(* IEC 61131-3 sources: plc-st-coding-agent/progress/evidence/f14_p1_20261111b/jobs/custom_deepseek-v4pro (part 2) *)

(* ---- self-hard-05.candidate_02.st ---- *)
FUNCTION_BLOCK FB
VAR_INPUT
    runRequest : BOOL;
    flameOK : BOOL;
    o2Valid : BOOL;
    o2PV : REAL;
    baseAir : REAL;
    resetBtn : BOOL;
END_VAR
VAR_OUTPUT
    fuelPermit : BOOL;
    trimEnable : BOOL;
    airTrim : REAL;
    airCommand : REAL;
    tripLatched : BOOL;
    o2Fault : BOOL;
END_VAR
VAR
    tripState : BOOL := FALSE;   (* internal trip memory *)
    prevReset : BOOL := FALSE;   (* previous cycle reset button state *)
    resetRising : BOOL;          (* reset rising edge flag *)
    rawTrim : REAL;              (* unclamped oxygen trim *)
END_VAR
BEGIN
    (* 1. Analyzer fault detection *)
    o2Fault := (NOT o2Valid) OR (o2PV < 0.0) OR (o2PV > 21.0);

    (* 2. Reset button rising edge detection *)
    resetRising := resetBtn AND (NOT prevReset);

    (* 3. Trip state update (immediate set, self-holding with edge-clear) *)
    IF (runRequest AND (NOT flameOK)) THEN
        tripState := TRUE;
    ELSIF (tripState AND resetRising AND (NOT runRequest) AND (NOT flameOK)) THEN
        tripState := FALSE;
    END_IF;

    (* 4. Output latched trip *)
    tripLatched := tripState;

    (* 5. Fuel permit *)
    fuelPermit := runRequest AND flameOK AND (NOT tripLatched);

    (* 6. Oxygen trim enable *)
    trimEnable := fuelPermit AND (NOT o2Fault);

    (* 7. Oxygen trim calculation *)
    IF trimEnable THEN
        rawTrim := 2.0 * (2.0 - o2PV);
        IF rawTrim < -10.0 THEN
            airTrim := -10.0;
        ELSIF rawTrim > 10.0 THEN
            airTrim := 10.0;
        ELSE
            airTrim := rawTrim;
        END_IF;
    ELSE
        airTrim := 0.0;
    END_IF;

    (* 8. Air command calculation *)
    IF fuelPermit THEN
        airCommand := baseAir + airTrim;
        IF airCommand < 0.0 THEN
            airCommand := 0.0;
        ELSIF airCommand > 100.0 THEN
            airCommand := 100.0;
        END_IF;
    ELSE
        airCommand := 0.0;
    END_IF;

    (* 9. Store reset button state for next cycle edge detection *)
    prevReset := resetBtn;
END_FUNCTION_BLOCK

(* ---- self-hard-06.candidate_01.st ---- *)
FUNCTION_BLOCK FB
VAR_INPUT
    runRequest : BOOL;
    pressure : REAL;
    pressureValid : BOOL;
    fuelFlow : REAL;
    steamFlow : REAL;
    outletCmd : INT;
    outletFeedback : INT;
    resetBtn : BOOL;
END_VAR
VAR_OUTPUT
    tripLatched : BOOL;
    fuelPermit : BOOL;
    currentCauseMask : WORD;
    latchedCauseMask : WORD;
    diagnosticActive : BOOL;
END_VAR
VAR
    stallCount : INT := 0;          (* 连续卡滞计数 *)
    prevResetBtn : BOOL := FALSE;   (* 上一周期复位按钮 *)
    risingReset : BOOL;
    condStall : BOOL;
    newTripLatched : BOOL;
END_VAR

(* 复位按钮上升沿检测 *)
risingReset := resetBtn AND NOT prevResetBtn;

(* 计算本拍诊断线索 currentCauseMask *)
currentCauseMask := 0;

IF NOT runRequest THEN
    currentCauseMask := 0;
    stallCount := 0;
ELSIF NOT pressureValid THEN
    currentCauseMask := 1;          (* bit0: 变送器失效 *)
    stallCount := 0;
ELSE
    (* runRequest AND pressureValid *)
    IF pressure < 4500.0 THEN
        currentCauseMask := 0;
        stallCount := 0;
    ELSE
        (* 超压工况: pressure >= 4500.0 *)
        condStall := (outletCmd >= 50) AND (outletFeedback <= 10);
        IF condStall THEN
            stallCount := stallCount + 1;
        ELSE
            stallCount := 0;
        END_IF

        (* bit1: 减温减压阀卡滞，连续3拍 *)
        IF stallCount >= 3 THEN
            currentCauseMask := currentCauseMask OR 16#0002;
        END_IF

        (* bit2: 燃烧过剩 *)
        IF (fuelFlow >= 4.0) AND (steamFlow <= 10.0) THEN
            currentCauseMask := currentCauseMask OR 16#0004;
        END_IF

        (* bit3: 未定位 *)
        IF currentCauseMask = 0 THEN
            currentCauseMask := 16#0008;
        END_IF
    END_IF
END_IF

(* 计算新的跳闸锁存状态 *)
newTripLatched := (runRequest AND (NOT pressureValid OR pressure >= 4500.0))
                  OR (tripLatched AND NOT (risingReset AND NOT runRequest AND pressureValid AND pressure <= 4200.0));

(* 更新跳闸期间线索累积足迹 *)
IF newTripLatched THEN
    latchedCauseMask := (latchedCauseMask OR currentCauseMask) AND 16#000F;
ELSE
    latchedCauseMask := 0;
END_IF

(* 输出更新 *)
tripLatched := newTripLatched;
fuelPermit := runRequest AND NOT newTripLatched;
diagnosticActive := (currentCauseMask <> 0);

(* 保存本拍 resetBtn 供下周期上升沿检测 *)
prevResetBtn := resetBtn;

(* ---- self-hard-06.candidate_02.st ---- *)
FUNCTION_BLOCK FB
VAR_INPUT
    runRequest : BOOL;
    pressure : REAL;
    pressureValid : BOOL;
    fuelFlow : REAL;
    steamFlow : REAL;
    outletCmd : INT;
    outletFeedback : INT;
    resetBtn : BOOL;
END_VAR
VAR_OUTPUT
    tripLatched : BOOL;
    fuelPermit : BOOL;
    currentCauseMask : WORD;
    latchedCauseMask : WORD;
    diagnosticActive : BOOL;
END_VAR
VAR
    stallCount : INT := 0;          (* 连续卡滞计数 *)
    prevResetBtn : BOOL := FALSE;   (* 上一周期复位按钮 *)
    risingReset : BOOL;
    condStall : BOOL;
    newTripLatched : BOOL;
END_VAR

(* 复位按钮上升沿检测 *)
risingReset := resetBtn AND NOT prevResetBtn;

(* 计算本拍诊断线索 currentCauseMask *)
currentCauseMask := 0;

IF NOT runRequest THEN
    currentCauseMask := 0;
    stallCount := 0;
ELSIF NOT pressureValid THEN
    currentCauseMask := 1;          (* bit0: 变送器失效 *)
    stallCount := 0;
ELSE
    (* runRequest AND pressureValid *)
    IF pressure < 4500.0 THEN
        currentCauseMask := 0;
        stallCount := 0;
    ELSE
        (* 超压工况: pressure >= 4500.0 *)
        condStall := (outletCmd >= 50) AND (outletFeedback <= 10);
        IF condStall THEN
            stallCount := stallCount + 1;
        ELSE
            stallCount := 0;
        END_IF

        (* bit1: 减温减压阀卡滞，连续3拍 *)
        IF stallCount >= 3 THEN
            currentCauseMask := currentCauseMask OR 16#0002;
        END_IF

        (* bit2: 燃烧过剩 *)
        IF (fuelFlow >= 4.0) AND (steamFlow <= 10.0) THEN
            currentCauseMask := currentCauseMask OR 16#0004;
        END_IF

        (* bit3: 未定位 *)
        IF currentCauseMask = 0 THEN
            currentCauseMask := 16#0008;
        END_IF
    END_IF
END_IF

(* 计算新的跳闸锁存状态 *)
newTripLatched := (runRequest AND (NOT pressureValid OR pressure >= 4500.0))
                  OR (tripLatched AND NOT (risingReset AND NOT runRequest AND pressureValid AND pressure <= 4200.0));

(* 更新跳闸期间线索累积足迹 *)
IF newTripLatched THEN
    latchedCauseMask := (latchedCauseMask OR currentCauseMask) AND 16#000F;
ELSE
    latchedCauseMask := 0;
END_IF

(* 输出更新 *)
tripLatched := newTripLatched;
fuelPermit := runRequest AND NOT newTripLatched;
diagnosticActive := (currentCauseMask <> 0);

(* 保存本拍 resetBtn 供下周期上升沿检测 *)
prevResetBtn := resetBtn;

END_FUNCTION_BLOCK

(* ---- self-medium-01.candidate_01.st ---- *)
TYPE ST_Recipe :
STRUCT
    recipeID : INT;
    totalRatio : REAL;
    temperature : REAL;
END_STRUCT
END_TYPE

FUNCTION_BLOCK FB
VAR_INPUT
    recipe : ARRAY[1..8] OF ST_Recipe;
    selSlot : INT;
    loadCmd : BOOL;
    running : BOOL;
END_VAR
VAR_OUTPUT
    valid : BOOL := FALSE;
    loadedID : INT := 0;
END_VAR
VAR
    prev_loadCmd : BOOL := FALSE;
END_VAR

// 仅在未生产且检测到 loadCmd 上升沿时执行装载校验
IF NOT running THEN
    IF loadCmd AND NOT prev_loadCmd THEN
        // 下标越界保护：先判断合法范围，避免访问数组外
        IF selSlot >= 1 AND selSlot <= 8 THEN
            // 校验：槽非空、总配比 [99.0, 101.0]、温度 [30.0, 180.0]
            IF recipe[selSlot].recipeID <> 0
               AND recipe[selSlot].totalRatio >= 99.0
               AND recipe[selSlot].totalRatio <= 101.0
               AND recipe[selSlot].temperature >= 30.0
               AND recipe[selSlot].temperature <= 180.0 THEN
                valid := TRUE;
                loadedID := recipe[selSlot].recipeID;
            ELSE
                valid := FALSE;
                loadedID := 0;
            END_IF
        ELSE
            valid := FALSE;
            loadedID := 0;
        END_IF
    END_IF
    // 无上升沿时，valid 和 loadedID 保持不变
END_IF
// running 为 TRUE 时，valid 和 loadedID 保持不变

// 更新上一周期命令状态，用于上升沿检测
prev_loadCmd := loadCmd;

END_FUNCTION_BLOCK

(* ---- self-medium-02.candidate_01.st ---- *)
FUNCTION_BLOCK FB
VAR_INPUT
    enable : BOOL;
    rawValue : REAL;
END_VAR
VAR_OUTPUT
    filteredValue : REAL;
    windowFull : BOOL;
    sampleCount : INT;
END_VAR
VAR
    buffer : ARRAY[0..7] OF REAL;
    count : INT := 0;
    sum : REAL;
    i : INT;
END_VAR

IF enable THEN
    // 更新缓冲区
    IF count < 8 THEN
        buffer[count] := rawValue;
        count := count + 1;
    ELSE
        // 满窗，FIFO左移
        FOR i := 0 TO 6 DO
            buffer[i] := buffer[i+1];
        END_FOR;
        buffer[7] := rawValue;
    END_IF;

    // 计算平均值
    sum := 0.0;
    FOR i := 0 TO count-1 DO
        sum := sum + buffer[i];
    END_FOR;
    filteredValue := sum / INT_TO_REAL(count);
ELSE
    // 停用：清空计数，保持filteredValue
    count := 0;
END_IF;

// 更新输出计数和满标志
sampleCount := count;
windowFull := (count = 8);

(* ---- self-medium-02.candidate_02.st ---- *)
FUNCTION_BLOCK FB
VAR_INPUT
    enable : BOOL;
    rawValue : REAL;
END_VAR
VAR_OUTPUT
    filteredValue : REAL;
    windowFull : BOOL;
    sampleCount : INT;
END_VAR
VAR
    buffer : ARRAY[0..7] OF REAL;
    count : INT := 0;
    sum : REAL;
    i : INT;
END_VAR

IF enable THEN
    // 更新缓冲区
    IF count < 8 THEN
        buffer[count] := rawValue;
        count := count + 1;
    ELSE
        // 满窗，FIFO左移
        FOR i := 0 TO 6 DO
            buffer[i] := buffer[i+1];
        END_FOR;
        buffer[7] := rawValue;
    END_IF;

    // 计算平均值
    sum := 0.0;
    FOR i := 0 TO count-1 DO
        sum := sum + buffer[i];
    END_FOR;
    filteredValue := sum / INT_TO_REAL(count);
ELSE
    // 停用：清空计数，保持filteredValue
    count := 0;
END_IF;

// 更新输出计数和满标志
sampleCount := count;
windowFull := (count = 8);

END_FUNCTION_BLOCK

(* ---- self-medium-03.candidate_01.st ---- *)
FUNCTION_BLOCK FB
VAR_INPUT
    openBtn : BOOL;
    closeBtn : BOOL;
    openLimit : BOOL;
    closeLimit : BOOL;
    obstacle : BOOL;
END_VAR
VAR_OUTPUT
    motorUp : BOOL;
    motorDown : BOOL;
    errorFlag : BOOL;
END_VAR
VAR
    prevOpenBtn : BOOL := FALSE;
    prevCloseBtn : BOOL := FALSE;
    prevBoth : BOOL := FALSE;
    prevMotorUp : BOOL := FALSE;
    prevMotorDown : BOOL := FALSE;
    prevErrorFlag : BOOL := FALSE;
    risingOpen : BOOL := FALSE;
    risingClose : BOOL := FALSE;
    currentBoth : BOOL := FALSE;
    risingBoth : BOOL := FALSE;
    state : INT := 0; (* 0:IDLE, 1:OPENING, 2:CLOSING, 3:FAULT *)
END_VAR

// 边沿检测
risingOpen := openBtn AND NOT prevOpenBtn;
risingClose := closeBtn AND NOT prevCloseBtn;
currentBoth := openBtn AND closeBtn;
risingBoth := currentBoth AND NOT prevBoth;

// 输出计算
motorUp := NOT obstacle AND NOT openLimit AND (prevMotorUp OR (NOT prevMotorUp AND NOT prevMotorDown AND NOT prevErrorFlag AND risingOpen AND NOT closeBtn));

motorDown := NOT obstacle AND NOT closeLimit AND (prevMotorDown OR (NOT prevMotorUp AND NOT prevMotorDown AND NOT prevErrorFlag AND risingClose AND NOT openBtn));

errorFlag := obstacle OR (prevErrorFlag AND NOT risingBoth);

// 状态更新
IF errorFlag THEN
    state := 3; // FAULT
ELSIF motorUp THEN
    state := 1; // OPENING
ELSIF motorDown THEN
    state := 2; // CLOSING
ELSE
    state := 0; // IDLE
END_IF;

// 更新 prev 变量
prevOpenBtn := openBtn;
prevCloseBtn := closeBtn;
prevBoth := currentBoth;
prevMotorUp := motorUp;
prevMotorDown := motorDown;
prevErrorFlag := errorFlag;

(* ---- self-medium-03.candidate_02.st ---- *)
FUNCTION_BLOCK FB
VAR_INPUT
    openBtn : BOOL;
    closeBtn : BOOL;
    openLimit : BOOL;
    closeLimit : BOOL;
    obstacle : BOOL;
END_VAR
VAR_OUTPUT
    motorUp : BOOL;
    motorDown : BOOL;
    errorFlag : BOOL;
END_VAR
VAR
    prevOpenBtn : BOOL := FALSE;
    prevCloseBtn : BOOL := FALSE;
    prevBoth : BOOL := FALSE;
    prevMotorUp : BOOL := FALSE;
    prevMotorDown : BOOL := FALSE;
    prevErrorFlag : BOOL := FALSE;
    risingOpen : BOOL := FALSE;
    risingClose : BOOL := FALSE;
    currentBoth : BOOL := FALSE;
    risingBoth : BOOL := FALSE;
    state : INT := 0;
END_VAR

// 边沿检测
risingOpen := openBtn AND NOT prevOpenBtn;
risingClose := closeBtn AND NOT prevCloseBtn;
currentBoth := openBtn AND closeBtn;
risingBoth := currentBoth AND NOT prevBoth;

// 输出计算
motorUp := NOT obstacle AND NOT openLimit AND (prevMotorUp OR (NOT prevMotorUp AND NOT prevMotorDown AND NOT prevErrorFlag AND risingOpen AND NOT closeBtn));

motorDown := NOT obstacle AND NOT closeLimit AND (prevMotorDown OR (NOT prevMotorUp AND NOT prevMotorDown AND NOT prevErrorFlag AND risingClose AND NOT openBtn));

errorFlag := obstacle OR (prevErrorFlag AND NOT risingBoth);

// 状态更新
IF errorFlag THEN
    state := 3; // FAULT
ELSIF motorUp THEN
    state := 1; // OPENING
ELSIF motorDown THEN
    state := 2; // CLOSING
ELSE
    state := 0; // IDLE
END_IF;

// 更新 prev 变量
prevOpenBtn := openBtn;
prevCloseBtn := closeBtn;
prevBoth := currentBoth;
prevMotorUp := motorUp;
prevMotorDown := motorDown;
prevErrorFlag := errorFlag;

END_FUNCTION_BLOCK

(* ---- self-medium-04.candidate_01.st ---- *)
FUNCTION_BLOCK FB
VAR_INPUT
    startBtn : BOOL;      (* 启动按钮，上升沿有效 *)
    resetBtn : BOOL;      (* 复位按钮，上升沿有效 *)
    doneSensor : BOOL;    (* 满瓶检测传感器 *)
    targetVol : REAL;     (* 目标灌装体积 mL *)
    flowVol : REAL;       (* 本周期累计流量增量 mL *)
END_VAR
VAR_OUTPUT
    valveOpen : BOOL;     (* 灌装阀开命令 *)
    fillsToday : INT;     (* 今日完成瓶数 *)
END_VAR
VAR
    prevStartBtn : BOOL := FALSE;   (* 上一周期启动按钮状态 *)
    prevResetBtn : BOOL := FALSE;   (* 上一周期复位按钮状态 *)
    accumVol : REAL := 0.0;         (* 本瓶累计灌装体积 *)
    pendingConfirm : BOOL := FALSE; (* 是否待确认 *)
    prevValveOpen : BOOL := FALSE;  (* 上一周期阀门状态 *)
END_VAR

    (* 保存上一周期阀门输出状态 *)
    prevValveOpen := valveOpen;

    (* 检测复位按钮上升沿，优先处理 *)
    IF (resetBtn AND NOT prevResetBtn) THEN
        (* 复位：清零计数、累计体积，关阀，清除待确认 *)
        valveOpen := FALSE;
        fillsToday := 0;
        accumVol := 0.0;
        pendingConfirm := FALSE;
    ELSE
        (* 非复位周期 *)

        (* 处理启动按钮上升沿（仅在阀门关闭时：空闲或等待确认） *)
        IF (startBtn AND NOT prevStartBtn) AND (NOT prevValveOpen) THEN
            (* 开始新瓶：清零本瓶累计，开阀，取消上一瓶待确认 *)
            accumVol := 0.0;
            pendingConfirm := FALSE;
            valveOpen := TRUE;
        END_IF;

        (* 正在灌装：累加本拍流量，检查是否达到目标 *)
        IF valveOpen THEN
            accumVol := accumVol + flowVol;
            IF accumVol >= targetVol THEN
                valveOpen := FALSE;
                pendingConfirm := TRUE;
            END_IF;
        END_IF;

        (* 处理确认：有待确认且传感器为真，则计数 *)
        IF pendingConfirm AND doneSensor THEN
            IF fillsToday < 32767 THEN
                fillsToday := fillsToday + 1;
            END_IF;
            pendingConfirm := FALSE;
        END_IF;
    END_IF;

    (* 更新按钮前一周期状态 *)
    prevStartBtn := startBtn;
    prevResetBtn := resetBtn;

END_FUNCTION_BLOCK

(* ---- self-medium-05.candidate_01.st ---- *)
FUNCTION_BLOCK FB
VAR_INPUT
    enable : BOOL;
    resetBtn : BOOL;
    scanSeconds : LREAL;
    steamFlow : LREAL;
    fuelFlow : LREAL;
    steamTemp : LREAL;
    steamPressure : LREAL;
END_VAR
VAR_OUTPUT
    qualified : BOOL;
    dataFault : BOOL;
    qualifiedTon : LREAL;
    fuelTon : LREAL;
    revenue : LREAL;
    cost : LREAL;
    netProfit : LREAL;
END_VAR
VAR
    prevReset : BOOL := FALSE;
    qAcc : LREAL := 0.0;
    fAcc : LREAL := 0.0;
END_VAR

qualified := (steamTemp >= 447.0) AND (steamTemp <= 453.0) AND (steamPressure >= 3750.0) AND (steamPressure <= 3850.0);

dataFault := (scanSeconds <= 0.0) OR (scanSeconds > 10.0) OR (steamFlow < 0.0) OR (steamFlow > 90.0) OR (fuelFlow < 0.0) OR (fuelFlow > 6.0);

IF resetBtn AND NOT prevReset THEN
    qAcc := 0.0;
    fAcc := 0.0;
ELSE
    IF enable AND NOT dataFault THEN
        fAcc := fAcc + (fuelFlow * scanSeconds / 1000.0);
        IF qualified THEN
            qAcc := qAcc + (steamFlow * scanSeconds / 1000.0);
        END_IF;
    END_IF;
END_IF;

qualifiedTon := qAcc;
fuelTon := fAcc;
revenue := qAcc * 280.0;
cost := fAcc * 1500.0;
netProfit := revenue - cost;

prevReset := resetBtn;
END_FUNCTION_BLOCK

(* ---- self-medium-06.candidate_01.st ---- *)
FUNCTION_BLOCK FB
VAR_INPUT
    enable : BOOL;
    resetBtn : BOOL;
    sensorValid : BOOL;
    setpoint : REAL;
    temperature : REAL;
    scanSeconds : REAL;
    bias : REAL;
END_VAR
VAR_OUTPUT
    power : REAL;
    correction : REAL;
    fault : BOOL;
END_VAR
VAR
    ePrev : REAL;
    histValid : BOOL;
    lastResetBtn : BOOL;
END_VAR
VAR_TEMP
    e : REAL;
    de : REAL;
    x : REAL;
    y : REAL;
    resetRising : BOOL;
END_VAR

BEGIN
    -- 计算误差
    e := setpoint - temperature;

    -- 计算故障
    fault := NOT sensorValid OR (scanSeconds <= 0.0) OR (scanSeconds > 10.0);

    -- 检测复位上升沿
    resetRising := resetBtn AND NOT lastResetBtn;

    IF (NOT enable OR fault OR resetRising) THEN
        -- 故障、停用或复位上升沿：输出归零，清除历史
        power := 0.0;
        correction := 0.0;
        ePrev := 0.0;
        histValid := FALSE;
    ELSE
        -- 正常模糊计算
        IF histValid THEN
            de := (e - ePrev) / scanSeconds;
        ELSE
            de := 0.0;  -- 首拍或历史被清除后恢复首拍
        END_IF;

        x := LIMIT(-1.0, e / 10.0, 1.0);
        y := LIMIT(-1.0, de / 2.0, 1.0);

        -- 九规则重心法等价于 20*x + 10*y
        correction := 20.0 * x + 10.0 * y;

        power := LIMIT(0.0, bias + correction, 100.0);

        ePrev := e;
        histValid := TRUE;
    END_IF;

    -- 更新上一周期复位按钮状态
    lastResetBtn := resetBtn;
END_FUNCTION_BLOCK

(* ---- self-medium-06.candidate_02.st ---- *)
FUNCTION_BLOCK FB
VAR_INPUT
    enable : BOOL;
    resetBtn : BOOL;
    sensorValid : BOOL;
    setpoint : REAL;
    temperature : REAL;
    scanSeconds : REAL;
    bias : REAL;
END_VAR
VAR_OUTPUT
    power : REAL;
    correction : REAL;
    fault : BOOL;
END_VAR
VAR
    ePrev : REAL;
    histValid : BOOL;
    lastResetBtn : BOOL;
END_VAR
VAR_TEMP
    e : REAL;
    de : REAL;
    x : REAL;
    y : REAL;
    resetRising : BOOL;
    tempPower : REAL;
END_VAR

BEGIN
    -- Compute error
    e := setpoint - temperature;

    -- Compute fault status
    fault := NOT sensorValid OR (scanSeconds <= 0.0) OR (scanSeconds > 10.0);

    -- Detect rising edge of reset button
    resetRising := resetBtn AND NOT lastResetBtn;

    IF (NOT enable OR fault OR resetRising) THEN
        -- Fault, disabled, or reset rising edge:
        -- Output zero and clear history
        power := 0.0;
        correction := 0.0;
        ePrev := 0.0;
        histValid := FALSE;
    ELSE
        -- Normal fuzzy calculation
        IF histValid THEN
            de := (e - ePrev) / scanSeconds;
        ELSE
            de := 0.0;  -- First cycle after start/reset/fault recovery
        END_IF;

        -- Clamp x to [-1, 1]
        x := e / 10.0;
        IF x < -1.0 THEN
            x := -1.0;
        ELSIF x > 1.0 THEN
            x := 1.0;
        END_IF;

        -- Clamp y to [-1, 1]
        y := de / 2.0;
        IF y < -1.0 THEN
            y := -1.0;
        ELSIF y > 1.0 THEN
            y := 1.0;
        END_IF;

        -- Nine-rule centroid equivalent: 20*x + 10*y
        correction := 20.0 * x + 10.0 * y;

        -- Clamp power to [0, 100]
        tempPower := bias + correction;
        IF tempPower < 0.0 THEN
            power := 0.0;
        ELSIF tempPower > 100.0 THEN
            power := 100.0;
        ELSE
            power := tempPower;
        END_IF;

        -- Update history
        ePrev := e;
        histValid := TRUE;
    END_IF;

    -- Store current reset button state for next cycle edge detection
    lastResetBtn := resetBtn;
END_FUNCTION_BLOCK

(* ---- public-easy-01.candidate_01.st ---- *)
PROGRAM AutomatedFillingLine
VAR_INPUT
    bottleSensor         : BOOL;  // Bottle detection sensor
    cleaningConfirmButton : BOOL; // Cleaning completion confirmation
    fillingConfirmButton  : BOOL; // Filling completion confirmation
    cappingConfirmButton  : BOOL; // Capping completion confirmation
    packingConfirmButton  : BOOL; // Packaging completion confirmation
    finishedButton        : BOOL; // Bottle pickup confirmation
END_VAR
VAR_OUTPUT
    Pump_Motor        : BOOL; // Cleaning pump motor
    Filling_Valve     : BOOL; // Filling valve
    Capping_Machine   : BOOL; // Capping machine
    Packing_Machine   : BOOL; // Packing machine
    Completion_Light  : BOOL; // Packaging completion indicator
END_VAR
VAR
    state    : INT := 0; // 0=Idle, 1=Cleaning, 2=Filling, 3=Capping, 4=Packing, 5=Complete
    rBottle  : R_TRIG;
    rClean   : R_TRIG;
    rFill    : R_TRIG;
    rCap     : R_TRIG;
    rPack    : R_TRIG;
    rFinish  : R_TRIG;
END_VAR

// Edge detection for all digital signals
rBottle(CLK := bottleSensor);
rClean(CLK := cleaningConfirmButton);
rFill(CLK := fillingConfirmButton);
rCap(CLK := cappingConfirmButton);
rPack(CLK := packingConfirmButton);
rFinish(CLK := finishedButton);

CASE state OF
    // Idle: wait for bottle sensor
    0:
        Pump_Motor := FALSE;
        Filling_Valve := FALSE;
        Capping_Machine := FALSE;
        Packing_Machine := FALSE;
        Completion_Light := FALSE;

        IF rBottle.Q THEN
            state := 1;              // Start cleaning
            Pump_Motor := TRUE;
        END_IF;

    // Cleaning: run pump until operator confirms
    1:
        Pump_Motor := TRUE;
        Filling_Valve := FALSE;
        Capping_Machine := FALSE;
        Packing_Machine := FALSE;
        Completion_Light := FALSE;

        IF rClean.Q THEN
            state := 2;              // Cleaning done, start filling
            Pump_Motor := FALSE;
            Filling_Valve := TRUE;
        END_IF;

    // Filling: open valve until operator confirms
    2:
        Pump_Motor := FALSE;
        Filling_Valve := TRUE;
        Capping_Machine := FALSE;
        Packing_Machine := FALSE;
        Completion_Light := FALSE;

        IF rFill.Q THEN
            state := 3;              // Filling done, start capping
            Filling_Valve := FALSE;
            Capping_Machine := TRUE;
        END_IF;

    // Capping: run capping machine until operator confirms
    3:
        Pump_Motor := FALSE;
        Filling_Valve := FALSE;
        Capping_Machine := TRUE;
        Packing_Machine := FALSE;
        Completion_Light := FALSE;

        IF rCap.Q THEN
            state := 4;              // Capping done, start packing
            Capping_Machine := FALSE;
            Packing_Machine := TRUE;
        END_IF;

    // Packing: run packing machine until operator confirms
    4:
        Pump_Motor := FALSE;
        Filling_Valve := FALSE;
        Capping_Machine := FALSE;
        Packing_Machine := TRUE;
        Completion_Light := FALSE;

        IF rPack.Q THEN
            state := 5;              // Packing done, light indicator
            Packing_Machine := FALSE;
            Completion_Light := TRUE;
        END_IF;

    // Complete: wait for operator to pick up bottle
    5:
        Pump_Motor := FALSE;
        Filling_Valve := FALSE;
        Capping_Machine := FALSE;
        Packing_Machine := FALSE;
        Completion_Light := TRUE;

        IF rFinish.Q THEN
            state := 0;              // Reset for next bottle
            Completion_Light := FALSE;
        END_IF;
END_CASE;

(* ---- public-easy-01.candidate_02.st ---- *)
PROGRAM AutomatedFillingLine
VAR_INPUT
    bottleSensor         : BOOL;  // Bottle detection sensor
    cleaningConfirmButton : BOOL; // Cleaning completion confirmation
    fillingConfirmButton  : BOOL; // Filling completion confirmation
    cappingConfirmButton  : BOOL; // Capping completion confirmation
    packingConfirmButton  : BOOL; // Packaging completion confirmation
    finishedButton        : BOOL; // Bottle pickup confirmation
END_VAR
VAR_OUTPUT
    Pump_Motor        : BOOL; // Cleaning pump motor
    Filling_Valve     : BOOL; // Filling valve
    Capping_Machine   : BOOL; // Capping machine
    Packing_Machine   : BOOL; // Packing machine
    Completion_Light  : BOOL; // Packaging completion indicator
END_VAR
VAR
    state    : INT := 0; // 0=Idle, 1=Cleaning, 2=Filling, 3=Capping, 4=Packing, 5=Complete
    rBottle  : R_TRIG;
    rClean   : R_TRIG;
    rFill    : R_TRIG;
    rCap     : R_TRIG;
    rPack    : R_TRIG;
    rFinish  : R_TRIG;
END_VAR

// Edge detection for all digital signals
rBottle(CLK := bottleSensor);
rClean(CLK := cleaningConfirmButton);
rFill(CLK := fillingConfirmButton);
rCap(CLK := cappingConfirmButton);
rPack(CLK := packingConfirmButton);
rFinish(CLK := finishedButton);

CASE state OF
    // Idle: wait for bottle sensor
    0:
        Pump_Motor := FALSE;
        Filling_Valve := FALSE;
        Capping_Machine := FALSE;
        Packing_Machine := FALSE;
        Completion_Light := FALSE;

        IF rBottle.Q THEN
            state := 1;              // Start cleaning
            Pump_Motor := TRUE;
        END_IF;

    // Cleaning: run pump until operator confirms
    1:
        Pump_Motor := TRUE;
        Filling_Valve := FALSE;
        Capping_Machine := FALSE;
        Packing_Machine := FALSE;
        Completion_Light := FALSE;

        IF rClean.Q THEN
            state := 2;              // Cleaning done, start filling
            Pump_Motor := FALSE;
            Filling_Valve := TRUE;
        END_IF;

    // Filling: open valve until operator confirms
    2:
        Pump_Motor := FALSE;
        Filling_Valve := TRUE;
        Capping_Machine := FALSE;
        Packing_Machine := FALSE;
        Completion_Light := FALSE;

        IF rFill.Q THEN
            state := 3;              // Filling done, start capping
            Filling_Valve := FALSE;
            Capping_Machine := TRUE;
        END_IF;

    // Capping: run capping machine until operator confirms
    3:
        Pump_Motor := FALSE;
        Filling_Valve := FALSE;
        Capping_Machine := TRUE;
        Packing_Machine := FALSE;
        Completion_Light := FALSE;

        IF rCap.Q THEN
            state := 4;              // Capping done, start packing
            Capping_Machine := FALSE;
            Packing_Machine := TRUE;
        END_IF;

    // Packing: run packing machine until operator confirms
    4:
        Pump_Motor := FALSE;
        Filling_Valve := FALSE;
        Capping_Machine := FALSE;
        Packing_Machine := TRUE;
        Completion_Light := FALSE;

        IF rPack.Q THEN
            state := 5;              // Packing done, light indicator
            Packing_Machine := FALSE;
            Completion_Light := TRUE;
        END_IF;

    // Complete: wait for operator to pick up bottle
    5:
        Pump_Motor := FALSE;
        Filling_Valve := FALSE;
        Capping_Machine := FALSE;
        Packing_Machine := FALSE;
        Completion_Light := TRUE;

        IF rFinish.Q THEN
            state := 0;              // Reset for next bottle
            Completion_Light := FALSE;
        END_IF;
END_CASE;

END_PROGRAM

(* ---- public-easy-04.candidate_01.st ---- *)
// Convert TIME inputs to LTIME for accumulation and comparison
CycleTime_LTIME := TIME_TO_LTIME(CycleTime);
DebounceTime_LTIME := TIME_TO_LTIME(DebounceTime);

// Viscosity debouncing
IF NOT VISCOSITY_OK THEN
    // Invalidate immediately on false
    ViscosityValid := FALSE;
    DebounceTimer := LTIME#0s;
ELSIF NOT ViscosityValid THEN
    // Only accumulate debounce time when emergency stop is not active
    IF PASTE_E_STOP_NC THEN
        DebounceTimer := DebounceTimer + CycleTime_LTIME;
    ELSE
        // Emergency stop clears any incomplete debounce timing
        DebounceTimer := LTIME#0s;
    END_IF;

    // Check if debounce time has been reached
    IF DebounceTimer >= DebounceTime_LTIME THEN
        ViscosityValid := TRUE;
        DebounceTimer := DebounceTime_LTIME; // Clamp to avoid overflow
    END_IF;
END_IF;

// Emergency stop priority: run output only when e-stop closed and viscosity valid
IF PASTE_E_STOP_NC AND ViscosityValid THEN
    VFD_RUN := TRUE;
ELSE
    VFD_RUN := FALSE;
END_IF;

// Accumulate runtime only while pump is running
IF VFD_RUN THEN
    PUMP_RUNTIME_ACC := PUMP_RUNTIME_ACC + CycleTime_LTIME;
END_IF;

// Maintenance due latching at 500 hours
IF NOT PUMP_MAINT_DUE AND (PUMP_RUNTIME_ACC >= LTIME#500h) THEN
    PUMP_MAINT_DUE := TRUE;
END_IF;

(* ---- public-hard-01.candidate_01.st ---- *)
PROGRAM MaterialProportioningControl
VAR_INPUT
    estop : BOOL;
    opeMode : BOOL;
    valveAStart : BOOL;
    valveBStart : BOOL;
    valveCStart : BOOL;
    valveDStart : BOOL;
    mixMotorStart : BOOL;
    autoStart : BOOL;
    processMode : BOOL;
    levelSensor : INT;
    mixMotorComplete : BOOL;
END_VAR
VAR_OUTPUT
    valveARun : BOOL;
    valveBRun : BOOL;
    valveCRun : BOOL;
    valveDRun : BOOL;
    mixMotorRun : BOOL;
END_VAR
VAR
    (* Previous states for edge detection *)
    prevValveAStart : BOOL;
    prevValveBStart : BOOL;
    prevValveCStart : BOOL;
    prevValveDStart : BOOL;
    prevMixMotorStart : BOOL;
    prevAutoStart : BOOL;
    prevMixMotorComplete : BOOL;

    (* Rising edge flags *)
    valveAStartRise : BOOL;
    valveBStartRise : BOOL;
    valveCStartRise : BOOL;
    valveDStartRise : BOOL;
    mixMotorStartRise : BOOL;
    autoStartRise : BOOL;
    mixMotorCompleteRise : BOOL;

    (* Automatic process state *)
    autoState : INT := 0;
    (* 0  - idle
       10 - filling A
       20 - filling B
       30 - filling C (only when processMode = TRUE)
       40 - mixing
       50 - discharging / process complete *)
END_VAR

(* --- Edge detection --- *)
valveAStartRise := valveAStart AND NOT prevValveAStart;
valveBStartRise := valveBStart AND NOT prevValveBStart;
valveCStartRise := valveCStart AND NOT prevValveCStart;
valveDStartRise := valveDStart AND NOT prevValveDStart;
mixMotorStartRise := mixMotorStart AND NOT prevMixMotorStart;
autoStartRise := autoStart AND NOT prevAutoStart;
mixMotorCompleteRise := mixMotorComplete AND NOT prevMixMotorComplete;

(* --- Emergency stop: stop everything immediately --- *)
IF NOT estop THEN
    valveARun := FALSE;
    valveBRun := FALSE;
    valveCRun := FALSE;
    valveDRun := FALSE;
    mixMotorRun := FALSE;
    autoState := 0;

(* --- Manual mode --- *)
ELSIF NOT opeMode THEN
    autoState := 0;

    IF valveAStartRise THEN
        valveARun := NOT valveARun;
    END_IF;

    IF valveBStartRise THEN
        valveBRun := NOT valveBRun;
    END_IF;

    IF valveCStartRise THEN
        valveCRun := NOT valveCRun;
    END_IF;

    IF valveDStartRise THEN
        valveDRun := NOT valveDRun;
    END_IF;

    IF mixMotorStartRise THEN
        mixMotorRun := NOT mixMotorRun;
    END_IF;

(* --- Automatic mode --- *)
ELSE
    (* Default all outputs off; the active state will turn on what is needed *)
    valveARun := FALSE;
    valveBRun := FALSE;
    valveCRun := FALSE;
    valveDRun := FALSE;
    mixMotorRun := FALSE;

    (* Start a new automatic process from idle or done state *)
    IF autoStartRise AND (autoState = 0 OR autoState = 50) THEN
        autoState := 10;
    END_IF;

    CASE autoState OF
        10: (* Filling with material A *)
            valveARun := TRUE;
            IF levelSensor >= 50 THEN
                autoState := 20;
            END_IF;

        20: (* Filling with material B *)
            valveBRun := TRUE;
            IF levelSensor >= 80 THEN
                IF processMode THEN
                    autoState := 30;
                ELSE
                    autoState := 40;
                END_IF;
            END_IF;

        30: (* Filling with material C, only processMode = TRUE *)
            valveCRun := TRUE;
            IF levelSensor >= 100 THEN
                autoState := 40;
            END_IF;

        40: (* Mixing *)
            mixMotorRun := TRUE;
            IF mixMotorCompleteRise THEN
                mixMotorRun := FALSE;
                autoState := 50;
            END_IF;

        50: (* Discharge through valve D, process complete *)
            valveDRun := TRUE;
    END_CASE;
END_IF;

(* --- Store current states for next scan --- *)
prevValveAStart := valveAStart;
prevValveBStart := valveBStart;
prevValveCStart := valveCStart;
prevValveDStart := valveDStart;
prevMixMotorStart := mixMotorStart;
prevAutoStart := autoStart;
prevMixMotorComplete := mixMotorComplete;

(* ---- public-hard-01.candidate_02.st ---- *)
PROGRAM MaterialProportioningControl
VAR_INPUT
    estop : BOOL;
    opeMode : BOOL;
    valveAStart : BOOL;
    valveBStart : BOOL;
    valveCStart : BOOL;
    valveDStart : BOOL;
    mixMotorStart : BOOL;
    autoStart : BOOL;
    processMode : BOOL;
    levelSensor : INT;
    mixMotorComplete : BOOL;
END_VAR
VAR_OUTPUT
    valveARun : BOOL;
    valveBRun : BOOL;
    valveCRun : BOOL;
    valveDRun : BOOL;
    mixMotorRun : BOOL;
END_VAR
VAR
    (* Previous states for edge detection *)
    prevValveAStart : BOOL;
    prevValveBStart : BOOL;
    prevValveCStart : BOOL;
    prevValveDStart : BOOL;
    prevMixMotorStart : BOOL;
    prevAutoStart : BOOL;
    prevMixMotorComplete : BOOL;

    (* Rising edge flags *)
    valveAStartRise : BOOL;
    valveBStartRise : BOOL;
    valveCStartRise : BOOL;
    valveDStartRise : BOOL;
    mixMotorStartRise : BOOL;
    autoStartRise : BOOL;
    mixMotorCompleteRise : BOOL;

    (* Automatic process state *)
    autoState : INT := 0;
    (* 0  - idle
       10 - filling A
       20 - filling B
       30 - filling C (only when processMode = TRUE)
       40 - mixing
       50 - discharging / process complete *)
END_VAR

(* --- Edge detection --- *)
valveAStartRise := valveAStart AND NOT prevValveAStart;
valveBStartRise := valveBStart AND NOT prevValveBStart;
valveCStartRise := valveCStart AND NOT prevValveCStart;
valveDStartRise := valveDStart AND NOT prevValveDStart;
mixMotorStartRise := mixMotorStart AND NOT prevMixMotorStart;
autoStartRise := autoStart AND NOT prevAutoStart;
mixMotorCompleteRise := mixMotorComplete AND NOT prevMixMotorComplete;

(* --- Emergency stop: stop everything immediately --- *)
IF NOT estop THEN
    valveARun := FALSE;
    valveBRun := FALSE;
    valveCRun := FALSE;
    valveDRun := FALSE;
    mixMotorRun := FALSE;
    autoState := 0;

(* --- Manual mode --- *)
ELSIF NOT opeMode THEN
    autoState := 0;

    IF valveAStartRise THEN
        valveARun := NOT valveARun;
    END_IF;

    IF valveBStartRise THEN
        valveBRun := NOT valveBRun;
    END_IF;

    IF valveCStartRise THEN
        valveCRun := NOT valveCRun;
    END_IF;

    IF valveDStartRise THEN
        valveDRun := NOT valveDRun;
    END_IF;

    IF mixMotorStartRise THEN
        mixMotorRun := NOT mixMotorRun;
    END_IF;

(* --- Automatic mode --- *)
ELSE
    (* Default all outputs off; the active state will turn on what is needed *)
    valveARun := FALSE;
    valveBRun := FALSE;
    valveCRun := FALSE;
    valveDRun := FALSE;
    mixMotorRun := FALSE;

    (* Start a new automatic process from idle or done state *)
    IF autoStartRise AND (autoState = 0 OR autoState = 50) THEN
        autoState := 10;
    END_IF;

    CASE autoState OF
        10: (* Filling with material A *)
            valveARun := TRUE;
            IF levelSensor >= 50 THEN
                autoState := 20;
            END_IF;

        20: (* Filling with material B *)
            valveBRun := TRUE;
            IF levelSensor >= 80 THEN
                IF processMode THEN
                    autoState := 30;
                ELSE
                    autoState := 40;
                END_IF;
            END_IF;

        30: (* Filling with material C, only processMode = TRUE *)
            valveCRun := TRUE;
            IF levelSensor >= 100 THEN
                autoState := 40;
            END_IF;

        40: (* Mixing *)
            mixMotorRun := TRUE;
            IF mixMotorCompleteRise THEN
                mixMotorRun := FALSE;
                autoState := 50;
            END_IF;

        50: (* Discharge through valve D, process complete *)
            valveDRun := TRUE;
    END_CASE;
END_IF;

(* --- Store current states for next scan --- *)
prevValveAStart := valveAStart;
prevValveBStart := valveBStart;
prevValveCStart := valveCStart;
prevValveDStart := valveDStart;
prevMixMotorStart := mixMotorStart;
prevAutoStart := autoStart;
prevMixMotorComplete := mixMotorComplete;

END_PROGRAM

(* ---- public-hard-05.candidate_01.st ---- *)
PROGRAM MechanicalArmControl
VAR_INPUT
    ManualMode: BOOL;
    SingleStepMode: BOOL;
    SingleCycleMode: BOOL;
    ContinuousMode: BOOL;
    EmergencyStop: BOOL;
    Start: BOOL;
    DownButton: BOOL;
    UpButton: BOOL;
    LeftButton: BOOL;
    RightButton: BOOL;
    GripButton: BOOL;
    ReleaseButton: BOOL;
    DownLimitSwitch: BOOL;
    UpLimitSwitch: BOOL;
    LeftLimitSwitch: BOOL;
    RightLimitSwitch: BOOL;
    GripLimitSwitch: BOOL;
    ReleaseLimitSwitch: BOOL;
END_VAR
VAR_OUTPUT
    MoveDown: BOOL;
    MoveUp: BOOL;
    MoveLeft: BOOL;
    MoveRight: BOOL;
    ActivateGrip: BOOL;
    ActivateRelease: BOOL;
END_VAR
VAR
    prevStart: BOOL := FALSE;
    startRising: BOOL;
    stepIndex: INT := 0;
    executing: BOOL := FALSE;
END_VAR

// Rising edge detection for Start button
startRising := Start AND NOT prevStart;
prevStart := Start;

IF NOT EmergencyStop THEN
    // Emergency stop active: stop all actions and reset automatic state
    executing := FALSE;
    stepIndex := 0;
ELSE
    // Normal operation
    IF ManualMode THEN
        // Manual mode: no automatic state; reset if switching from auto
        executing := FALSE;
        stepIndex := 0;
    ELSIF SingleStepMode THEN
        // Single step mode: one action per Start press
        IF startRising AND NOT executing THEN
            executing := TRUE;
        END_IF;
        IF executing THEN
            CASE stepIndex OF
                0: IF DownLimitSwitch THEN executing := FALSE; stepIndex := 1; END_IF
                1: IF GripLimitSwitch THEN executing := FALSE; stepIndex := 2; END_IF
                2: IF UpLimitSwitch THEN executing := FALSE; stepIndex := 3; END_IF
                3: IF RightLimitSwitch THEN executing := FALSE; stepIndex := 4; END_IF
                4: IF DownLimitSwitch THEN executing := FALSE; stepIndex := 5; END_IF
                5: IF ReleaseLimitSwitch THEN executing := FALSE; stepIndex := 6; END_IF
                6: IF UpLimitSwitch THEN executing := FALSE; stepIndex := 7; END_IF
                7: IF LeftLimitSwitch THEN executing := FALSE; stepIndex := 0; END_IF
            END_CASE;
        END_IF;
    ELSIF SingleCycleMode THEN
        // Single cycle mode: full cycle once per Start press
        IF startRising AND NOT executing THEN
            executing := TRUE;
            stepIndex := 0;
        END_IF;
        IF executing THEN
            CASE stepIndex OF
                0: IF DownLimitSwitch THEN stepIndex := 1; END_IF
                1: IF GripLimitSwitch THEN stepIndex := 2; END_IF
                2: IF UpLimitSwitch THEN stepIndex := 3; END_IF
                3: IF RightLimitSwitch THEN stepIndex := 4; END_IF
                4: IF DownLimitSwitch THEN stepIndex := 5; END_IF
                5: IF ReleaseLimitSwitch THEN stepIndex := 6; END_IF
                6: IF UpLimitSwitch THEN stepIndex := 7; END_IF
                7: IF LeftLimitSwitch THEN
                        executing := FALSE;
                        stepIndex := 0;
                    END_IF
            END_CASE;
        END_IF;
    ELSIF ContinuousMode THEN
        // Continuous mode: repeat cycles until stopped
        IF startRising AND NOT executing THEN
            executing := TRUE;
            stepIndex := 0;
        END_IF;
        IF executing THEN
            CASE stepIndex OF
                0: IF DownLimitSwitch THEN stepIndex := 1; END_IF
                1: IF GripLimitSwitch THEN stepIndex := 2; END_IF
                2: IF UpLimitSwitch THEN stepIndex := 3; END_IF
                3: IF RightLimitSwitch THEN stepIndex := 4; END_IF
                4: IF DownLimitSwitch THEN stepIndex := 5; END_IF
                5: IF ReleaseLimitSwitch THEN stepIndex := 6; END_IF
                6: IF UpLimitSwitch THEN stepIndex := 7; END_IF
                7: IF LeftLimitSwitch THEN stepIndex := 0; END_IF
            END_CASE;
        END_IF;
    ELSE
        // No valid mode selected
        executing := FALSE;
        stepIndex := 0;
    END_IF;
END_IF;

// Output assignment
MoveDown := FALSE;
MoveUp := FALSE;
MoveLeft := FALSE;
MoveRight := FALSE;
ActivateGrip := FALSE;
ActivateRelease := FALSE;

IF EmergencyStop THEN
    IF ManualMode THEN
        MoveDown := DownButton AND NOT DownLimitSwitch;
        MoveUp := UpButton AND NOT UpLimitSwitch;
        MoveLeft := LeftButton AND NOT LeftLimitSwitch;
        MoveRight := RightButton AND NOT RightLimitSwitch;
        ActivateGrip := GripButton AND NOT GripLimitSwitch;
        ActivateRelease := ReleaseButton AND NOT ReleaseLimitSwitch;
    ELSIF SingleStepMode OR SingleCycleMode OR ContinuousMode THEN
        IF executing THEN
            CASE stepIndex OF
                0: MoveDown := NOT DownLimitSwitch;
                1: ActivateGrip := NOT GripLimitSwitch;
                2: MoveUp := NOT UpLimitSwitch;
                3: MoveRight := NOT RightLimitSwitch;
                4: MoveDown := NOT DownLimitSwitch;
                5: ActivateRelease := NOT ReleaseLimitSwitch;
                6: MoveUp := NOT UpLimitSwitch;
                7: MoveLeft := NOT LeftLimitSwitch;
            END_CASE;
        END_IF;
    END_IF;
END_IF;

(* ---- public-hard-05.candidate_02.st ---- *)
PROGRAM MechanicalArmControl
VAR_INPUT
    ManualMode: BOOL;
    SingleStepMode: BOOL;
    SingleCycleMode: BOOL;
    ContinuousMode: BOOL;
    EmergencyStop: BOOL;
    Start: BOOL;
    DownButton: BOOL;
    UpButton: BOOL;
    LeftButton: BOOL;
    RightButton: BOOL;
    GripButton: BOOL;
    ReleaseButton: BOOL;
    DownLimitSwitch: BOOL;
    UpLimitSwitch: BOOL;
    LeftLimitSwitch: BOOL;
    RightLimitSwitch: BOOL;
    GripLimitSwitch: BOOL;
    ReleaseLimitSwitch: BOOL;
END_VAR
VAR_OUTPUT
    MoveDown: BOOL;
    MoveUp: BOOL;
    MoveLeft: BOOL;
    MoveRight: BOOL;
    ActivateGrip: BOOL;
    ActivateRelease: BOOL;
END_VAR
VAR
    prevStart: BOOL := FALSE;
    startRising: BOOL;
    stepIndex: INT := 0;
    executing: BOOL := FALSE;
END_VAR

// Rising edge detection for Start button
startRising := Start AND NOT prevStart;
prevStart := Start;

IF NOT EmergencyStop THEN
    // Emergency stop active: stop all actions and reset automatic state
    executing := FALSE;
    stepIndex := 0;
ELSE
    // Normal operation
    IF ManualMode THEN
        // Manual mode: no automatic state; reset if switching from auto
        executing := FALSE;
        stepIndex := 0;
    ELSIF SingleStepMode THEN
        // Single step mode: one action per Start press
        IF startRising AND NOT executing THEN
            executing := TRUE;
        END_IF;
        IF executing THEN
            CASE stepIndex OF
                0: IF DownLimitSwitch THEN executing := FALSE; stepIndex := 1; END_IF
                1: IF GripLimitSwitch THEN executing := FALSE; stepIndex := 2; END_IF
                2: IF UpLimitSwitch THEN executing := FALSE; stepIndex := 3; END_IF
                3: IF RightLimitSwitch THEN executing := FALSE; stepIndex := 4; END_IF
                4: IF DownLimitSwitch THEN executing := FALSE; stepIndex := 5; END_IF
                5: IF ReleaseLimitSwitch THEN executing := FALSE; stepIndex := 6; END_IF
                6: IF UpLimitSwitch THEN executing := FALSE; stepIndex := 7; END_IF
                7: IF LeftLimitSwitch THEN executing := FALSE; stepIndex := 0; END_IF
            END_CASE;
        END_IF;
    ELSIF SingleCycleMode THEN
        // Single cycle mode: full cycle once per Start press
        IF startRising AND NOT executing THEN
            executing := TRUE;
            stepIndex := 0;
        END_IF;
        IF executing THEN
            CASE stepIndex OF
                0: IF DownLimitSwitch THEN stepIndex := 1; END_IF
                1: IF GripLimitSwitch THEN stepIndex := 2; END_IF
                2: IF UpLimitSwitch THEN stepIndex := 3; END_IF
                3: IF RightLimitSwitch THEN stepIndex := 4; END_IF
                4: IF DownLimitSwitch THEN stepIndex := 5; END_IF
                5: IF ReleaseLimitSwitch THEN stepIndex := 6; END_IF
                6: IF UpLimitSwitch THEN stepIndex := 7; END_IF
                7: IF LeftLimitSwitch THEN
                        executing := FALSE;
                        stepIndex := 0;
                    END_IF
            END_CASE;
        END_IF;
    ELSIF ContinuousMode THEN
        // Continuous mode: repeat cycles until stopped
        IF startRising AND NOT executing THEN
            executing := TRUE;
            stepIndex := 0;
        END_IF;
        IF executing THEN
            CASE stepIndex OF
                0: IF DownLimitSwitch THEN stepIndex := 1; END_IF
                1: IF GripLimitSwitch THEN stepIndex := 2; END_IF
                2: IF UpLimitSwitch THEN stepIndex := 3; END_IF
                3: IF RightLimitSwitch THEN stepIndex := 4; END_IF
                4: IF DownLimitSwitch THEN stepIndex := 5; END_IF
                5: IF ReleaseLimitSwitch THEN stepIndex := 6; END_IF
                6: IF UpLimitSwitch THEN stepIndex := 7; END_IF
                7: IF LeftLimitSwitch THEN stepIndex := 0; END_IF
            END_CASE;
        END_IF;
    ELSE
        // No valid mode selected
        executing := FALSE;
        stepIndex := 0;
    END_IF;
END_IF;

// Output assignment
MoveDown := FALSE;
MoveUp := FALSE;
MoveLeft := FALSE;
MoveRight := FALSE;
ActivateGrip := FALSE;
ActivateRelease := FALSE;

IF EmergencyStop THEN
    IF ManualMode THEN
        MoveDown := DownButton AND NOT DownLimitSwitch;
        MoveUp := UpButton AND NOT UpLimitSwitch;
        MoveLeft := LeftButton AND NOT LeftLimitSwitch;
        MoveRight := RightButton AND NOT RightLimitSwitch;
        ActivateGrip := GripButton AND NOT GripLimitSwitch;
        ActivateRelease := ReleaseButton AND NOT ReleaseLimitSwitch;
    ELSIF SingleStepMode OR SingleCycleMode OR ContinuousMode THEN
        IF executing THEN
            CASE stepIndex OF
                0: MoveDown := NOT DownLimitSwitch;
                1: ActivateGrip := NOT GripLimitSwitch;
                2: MoveUp := NOT UpLimitSwitch;
                3: MoveRight := NOT RightLimitSwitch;
                4: MoveDown := NOT DownLimitSwitch;
                5: ActivateRelease := NOT ReleaseLimitSwitch;
                6: MoveUp := NOT UpLimitSwitch;
                7: MoveLeft := NOT LeftLimitSwitch;
            END_CASE;
        END_IF;
    END_IF;
END_IF;

END_PROGRAM
